// TIA Portal V19 export
// export: Created 2026-10-15T10:10:36.4706712Z, ExportSetting WithDefaults, DisplayName Totally Integrated Automation Portal, DisplayVersion V19, DisplayName TIA Portal Openness, DisplayVersion V19, DisplayName TIA Portal Version Control Interface, DisplayVersion V19, DisplayName STEP 7 Professional, DisplayVersion V19, DisplayName STEP 7 Safety, DisplayVersion V19, DisplayName WinCC Basic/Comfort/Advanced, DisplayVersion V19, DisplayName WinCC Unified, DisplayVersion V19
FUNCTION "ROLL_PB18" : Void   // FC26, SCL
{ S7_Optimized_Access := 'TRUE' }
VERSION : 0.1
// stored: AutoNumber true, IsIECCheckEnabled false, SetENOAutomatically false, UDAEnableTagReadback false
   VAR_TEMP
      r : Bool;
      a1 : Word;
      a2 : Word;
      activeDataBlock : Int;
      comparisonResults : Array[0..0] of Bool;
   END_VAR
BEGIN

   #r := FALSE;
   #a1 := W#16#0000;
   #a2 := W#16#0000;
   #activeDataBlock := 0;
   // PB18, STEP 5 network 1
   #r := ("ROLL_State".M[70, 2] OR "ROLL_State".M[70, 3] OR "ROLL_State".M[70, 4] OR "ROLL_State".M[70, 6] OR "ROLL_State".M[71, 0]);
   "ROLL_State".M[80, 5] := #r;
   // PB18, STEP 5 network 2
   #r := (((NOT "ROLL_IO".Output[112, 0]) AND (NOT "ROLL_IO".Output[112, 5]) AND "ROLL_State".M[20, 5]) OR ((NOT "ROLL_IO".Output[112, 0]) AND "ROLL_State".M[20, 3]) OR ((NOT "ROLL_IO".Output[112, 5]) AND "ROLL_State".M[20, 4]) OR ((NOT "ROLL_IO".Output[17, 7]) AND "ROLL_State".M[20, 7]) OR (("ROLL_State".M[20, 1] OR "ROLL_State".M[20, 2]) AND "ROLL_State".M[28, 4]));
   "ROLL_State".M[250, 0] := #r;
   // PB18, STEP 5 network 3
   #r := (((NOT "ROLL_IO".Output[113, 0]) AND "ROLL_State".M[22, 2]) OR ((NOT "ROLL_IO".Output[113, 1]) AND "ROLL_State".M[22, 3]) OR ((NOT "ROLL_IO".Output[113, 3]) AND "ROLL_IO".Output[113, 2] AND "ROLL_State".M[22, 4]) OR ((NOT "ROLL_IO".Output[113, 5]) AND "ROLL_IO".Output[113, 4] AND "ROLL_State".M[22, 5]) OR ("ROLL_IO".Input[124, 1] AND "ROLL_State".M[22, 0]) OR ("ROLL_IO".Input[124, 4] AND "ROLL_State".M[22, 1]) OR "ROLL_State".M[250, 0]);
   "ROLL_State".M[250, 0] := #r;
   // PB18, STEP 5 network 4
   #r := ((("ROLL_IO".Input[11, 1] OR "ROLL_IO".Input[11, 2] OR "ROLL_IO".Input[11, 3] OR "ROLL_IO".Input[11, 4] OR "ROLL_IO".Input[119, 6] OR "ROLL_IO".Input[119, 7] OR "ROLL_IO".Input[120, 0] OR "ROLL_IO".Input[120, 1]) AND "ROLL_IO".Input[12, 5] AND "ROLL_IO".Input[12, 7] AND "ROLL_State".M[23, 0]) OR (("ROLL_State".M[23, 2] OR "ROLL_State".M[23, 3]) AND "ROLL_State".M[63, 1]) OR ("ROLL_IO".Input[11, 0] AND "ROLL_IO".Input[11, 6] AND "ROLL_State".M[23, 1]) OR ("ROLL_IO".Input[11, 0] AND "ROLL_IO".Input[12, 1] AND "ROLL_IO".Input[12, 7] AND "ROLL_State".M[23, 0]) OR "ROLL_State".M[250, 0]);
   "ROLL_State".M[250, 0] := #r;
   // PB18, STEP 5 network 5
   #r := (((NOT "ROLL_IO".Output[20, 1]) AND "ROLL_State".M[24, 1]) OR "ROLL_State".M[250, 0]);
   "ROLL_State".M[250, 0] := #r;
   // PB18, STEP 5 network 6
   #r := ((((NOT "ROLL_IO".Output[20, 4]) OR (NOT "ROLL_IO".Output[22, 6])) AND "ROLL_State".M[25, 0]) OR "ROLL_State".M[250, 0]);
   "ROLL_State".M[250, 0] := #r;
   // PB18, STEP 5 network 7
   #r := (((NOT "ROLL_IO".Output[20, 5]) AND "ROLL_State".M[26, 6]) OR ((NOT "ROLL_IO".Output[20, 6]) AND "ROLL_State".M[26, 0]) OR ((NOT "ROLL_IO".Output[21, 4]) AND "ROLL_State".M[26, 5]) OR "ROLL_State".M[250, 0]);
   "ROLL_State".M[250, 0] := #r;
   // PB18, STEP 5 network 8
   #r := (((NOT "ROLL_IO".Output[20, 6]) AND "ROLL_State".M[27, 4]) OR ((NOT "ROLL_IO".Output[21, 6]) AND "ROLL_State".M[27, 5]) OR ((NOT "ROLL_State".M[80, 5]) AND "ROLL_State".M[27, 7]) OR "ROLL_State".M[250, 0]);
   "ROLL_State".M[250, 0] := #r;
   // PB18, STEP 5 network 9
   #r := ((("ROLL_IO".Output[112, 0] OR "ROLL_IO".Output[112, 5]) AND "ROLL_State".M[20, 5]) OR ("ROLL_IO".Output[112, 0] AND "ROLL_State".M[20, 3]) OR ("ROLL_IO".Output[112, 5] AND "ROLL_State".M[20, 4]) OR ("ROLL_IO".Output[17, 7] AND "ROLL_State".M[20, 7]));
   "ROLL_State".M[252, 0] := #r;
   // PB18, STEP 5 network 10
   #r := (((NOT "ROLL_IO".Output[113, 2]) AND "ROLL_IO".Output[113, 3] AND "ROLL_State".M[22, 4]) OR ((NOT "ROLL_IO".Output[113, 4]) AND "ROLL_IO".Output[113, 5] AND "ROLL_State".M[22, 5]) OR ("ROLL_IO".Output[113, 0] AND "ROLL_State".M[22, 2]) OR ("ROLL_IO".Output[113, 1] AND "ROLL_State".M[22, 3]) OR ("ROLL_IO".Input[124, 2] AND "ROLL_State".M[22, 0]) OR ("ROLL_IO".Input[124, 5] AND "ROLL_State".M[22, 1]) OR "ROLL_State".M[252, 0]);
   "ROLL_State".M[252, 0] := #r;
   // PB18, STEP 5 network 11
   #r := (((NOT "ROLL_IO".Output[23, 1]) AND ("ROLL_IO".Input[11, 1] OR "ROLL_IO".Input[11, 2] OR "ROLL_IO".Input[11, 3] OR "ROLL_IO".Input[11, 4] OR "ROLL_IO".Input[119, 6] OR "ROLL_IO".Input[119, 7] OR "ROLL_IO".Input[120, 0] OR "ROLL_IO".Input[120, 1]) AND "ROLL_IO".Input[11, 6] AND "ROLL_State".M[23, 1]) OR ((NOT "ROLL_State".M[63, 1]) AND ("ROLL_State".M[23, 2] OR "ROLL_State".M[23, 3])) OR (((("ROLL_IO".Input[11, 1] OR "ROLL_IO".Input[11, 2] OR "ROLL_IO".Input[11, 3] OR "ROLL_IO".Input[11, 4] OR "ROLL_IO".Input[119, 6] OR "ROLL_IO".Input[119, 7] OR "ROLL_IO".Input[120, 0] OR "ROLL_IO".Input[120, 1]) AND "ROLL_IO".Input[12, 1]) OR ("ROLL_IO".Input[11, 0] AND "ROLL_IO".Input[12, 5])) AND "ROLL_IO".Input[12, 7] AND "ROLL_State".M[23, 0]) OR "ROLL_State".M[252, 0]);
   "ROLL_State".M[252, 0] := #r;
   // PB18, STEP 5 network 12
   #r := (("ROLL_IO".Output[20, 1] AND "ROLL_State".M[24, 1]) OR "ROLL_State".M[252, 0]);
   "ROLL_State".M[252, 0] := #r;
   // PB18, STEP 5 network 13
   #r := (("ROLL_IO".Output[20, 4] AND "ROLL_IO".Output[22, 6] AND "ROLL_State".M[25, 0]) OR "ROLL_State".M[252, 0]);
   "ROLL_State".M[252, 0] := #r;
   // PB18, STEP 5 network 14
   #r := (("ROLL_IO".Output[20, 6] AND "ROLL_State".M[26, 0]) OR "ROLL_State".M[252, 0]);
   "ROLL_State".M[252, 0] := #r;
   // PB18, STEP 5 network 15
   #r := (("ROLL_IO".Output[20, 5] AND "ROLL_State".M[26, 6]) OR ("ROLL_IO".Output[20, 6] AND "ROLL_State".M[27, 4]) OR ("ROLL_IO".Output[21, 4] AND "ROLL_State".M[26, 5]) OR ("ROLL_IO".Output[21, 6] AND "ROLL_State".M[27, 5]) OR ("ROLL_State".M[27, 7] AND "ROLL_State".M[80, 5]) OR "ROLL_State".M[252, 0]);
   "ROLL_State".M[252, 0] := #r;
   // PB18, STEP 5 network 16
   RETURN;
END_FUNCTION
